// LS Electric XG5000 project: NewProject
// PLC LSPLC
// task ControlLoop: Kind=2 Priority=7 Device=250
// task Initialize: Kind=1 Priority=2
// task Trigger0: Kind=3 Priority=2 Device=M00000
// task Trigger1: Kind=3 Priority=3 Device=M00000 BitCondition=1
// task Trigger2: Kind=3 Priority=4 Device=M00000 BitCondition=2
// task Trigger3: Kind=3 Priority=5 Device=M00000 BitCondition=3
// task Trigger4: Kind=3 Priority=6 Device=M00000 BitCondition=4
// task Trigger5: Kind=3 Priority=7 Device=D000000 WordValue=65535
// task Trigger6: Kind=3 Priority=2 Device=D000000 WordValue=65535 WordCondition=1
// task Trigger7: Kind=3 Priority=3 Device=D000000 WordValue=65535 WordCondition=2
// task Trigger8: Kind=3 Priority=4 Device=D000000 WordValue=65535 WordCondition=3
// task Trigger9: Kind=3 Priority=5 Device=D000000 WordValue=65535 WordCondition=4

PROGRAM NewProgram (task: ControlLoop)

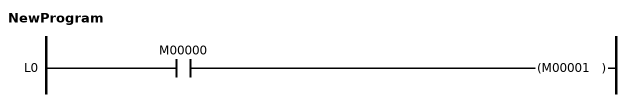
; L0
LOAD      M00000
OUT       M00001

PROGRAM ScanLoop (task: 스캔 프로그램)

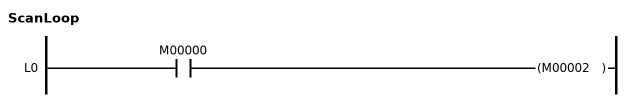
; L0
LOAD      M00000
OUT       M00002

PROGRAM Worker0 (task: Trigger0)

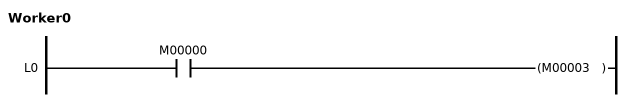
; L0
LOAD      M00000
OUT       M00003

PROGRAM Worker1 (task: Trigger1)

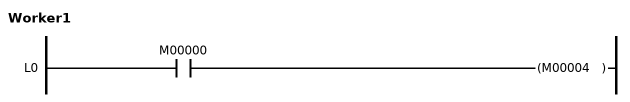
; L0
LOAD      M00000
OUT       M00004

PROGRAM Worker2 (task: Trigger2)

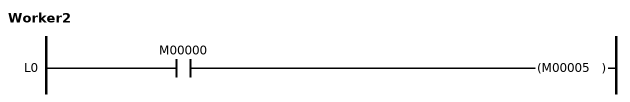
; L0
LOAD      M00000
OUT       M00005

PROGRAM Worker3 (task: Trigger3)

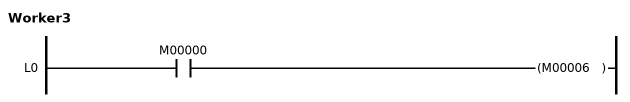
; L0
LOAD      M00000
OUT       M00006

PROGRAM Worker4 (task: Trigger4)

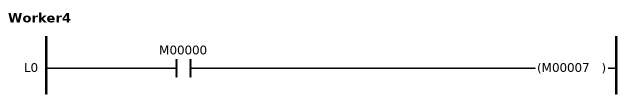
; L0
LOAD      M00000
OUT       M00007

PROGRAM Worker5 (task: Trigger5)

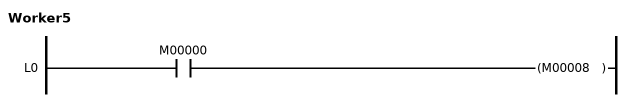
; L0
LOAD      M00000
OUT       M00008

PROGRAM Worker6 (task: Trigger6)

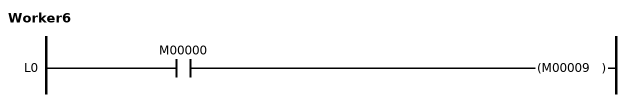
; L0
LOAD      M00000
OUT       M00009

PROGRAM Worker7 (task: Trigger7)

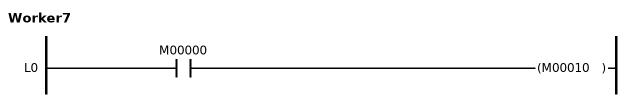
; L0
LOAD      M00000
OUT       M00010

PROGRAM Worker8 (task: Trigger8)

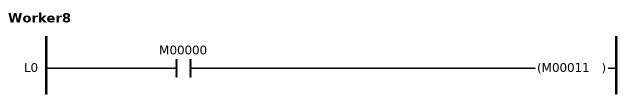
; L0
LOAD      M00000
OUT       M00011

PROGRAM Worker9 (task: Trigger9)

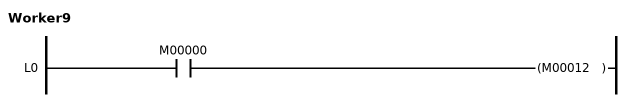
; L0
LOAD      M00000
OUT       M00012